Staubli VAL3: utCommon.dtx

public string sSource
public string sID
public string sPage
